Fanuc KAREL source: kc00001.KL

-- PROVISIONAL review KL for V1013-1; original PC SHA256 dba8aebd469e827f3fa26198d71ccb0bea972b9d083f9028c0a3483dfd4d9e0f
-- Incomplete behavior may be omitted. Consult companion uncertainty JSON. Do not deploy.
PROGRAM KC00001
%NOLOCKGROUP
BEGIN
  -- UNRESOLVED_PC offsets 5-14; opcodes 3F,75
  -- UNRESOLVED_PC offsets 19-28; opcodes 3F,75
  -- UNRESOLVED_PC offsets 33-71; opcodes 27,22,22,22,2A,22,2A,22,31
  -- UNRESOLVED_PC offsets 76-80; opcodes 7F
END KC00001
